(* IEC 61131-3 sources: plcassist-cli/packages/volt-lsp-iec/test-corpus/bakon-nano/Device/Plc Logic/Application/Library Manager/FloatingPointUtils, 43 files *)

(* ---- GVL.gvl ---- *)
VAR_GLOBAL
	EXP_MASK_REAL : UDINT := 16#7F800000;
	EXP_OFFSET_REAL : INT := 23;
	MANT_MASK_REAL : UDINT := 16#7FFFFF;
	RES_EXP_REAL : UINT := 16#FF;
	EXP_BIAS_REAL : INT := 127;
	NORM_MANT_REAL : UDINT := 16#800000;
	MAX_MANT_REAL : UDINT := 16#FFFFFF;
	MIN_EXP_REAL : INT := (INT#1 - (EXP_BIAS_REAL + EXP_OFFSET_REAL));
	MAX_EXP_REAL : INT := (UINT_TO_INT(RES_EXP_REAL) - ((INT#1 + EXP_BIAS_REAL) + EXP_OFFSET_REAL));
	EXP_MASK_LREAL : ULINT := 16#7FF0000000000000;
	EXP_OFFSET_LREAL : INT := 52;
	MANT_MASK_LREAL : ULINT := 16#FFFFFFFFFFFFF;
	RES_EXP_LREAL : UINT := 16#7FF;
	EXP_BIAS_LREAL : INT := 1023;
	NORM_MANT_LREAL : ULINT := 16#10000000000000;
	MAX_MANT_LREAL : ULINT := 16#1FFFFFFFFFFFFF;
	MIN_EXP_LREAL : INT := (INT#1 - (EXP_BIAS_LREAL + EXP_OFFSET_LREAL));
	MAX_EXP_LREAL : INT := (UINT_TO_INT(RES_EXP_LREAL) - ((INT#1 + EXP_BIAS_LREAL) + EXP_OFFSET_LREAL));
	STR_NAN : STRING(16) := 'NaN';
	STR_PINF : STRING(16) := '+Inf';
	STR_NINF : STRING(16) := '-Inf';
	LINT_MAX : LINT := 16#7FFFFFFFFFFFFFFF;
	INT_MAX : INT := 16#7FFF;
	INT_MIN : INT := -16#8000;
	DINT_MIN : DINT := -16#8000000;
	DINT_MAX : DINT := 16#7FFFFFFF;
END_VAR

(* ---- CEIL.fun ---- *)
FUNCTION CEIL : LREAL
VAR_INPUT
	F : LREAL;
END_VAR
END_FUNCTION

(* ---- CEILF.fun ---- *)
FUNCTION CEILF : REAL
VAR_INPUT
	F : REAL;
END_VAR
END_FUNCTION

(* ---- CHAREQCI.fun ---- *)
FUNCTION CHAREQCI : BOOL
VAR_INPUT
	C1 : BYTE;
	C2 : BYTE;
END_VAR
END_FUNCTION

(* ---- COMPOSELREAL.fun ---- *)
FUNCTION COMPOSELREAL : BOOL
VAR_INPUT
	LIM : LINT;
	IE : INT;
END_VAR
VAR_OUTPUT
	F : LREAL;
END_VAR
END_FUNCTION

(* ---- COMPOSELREALRAW.fun ---- *)
FUNCTION COMPOSELREALRAW : LREAL
VAR_INPUT
	BS : BOOL;
	UIE : UINT;
	ULIM : ULINT;
END_VAR
END_FUNCTION

(* ---- COMPOSEREAL.fun ---- *)
FUNCTION COMPOSEREAL : BOOL
VAR_INPUT
	DIM : DINT;
	IE : INT;
END_VAR
VAR_OUTPUT
	F : REAL;
END_VAR
END_FUNCTION

(* ---- COMPOSEREALRAW.fun ---- *)
FUNCTION COMPOSEREALRAW : REAL
VAR_INPUT
	BS : BOOL;
	UIE : UINT;
	UDIM : UDINT;
END_VAR
END_FUNCTION

(* ---- DESERIALIZEHEXREAL.fun ---- *)
FUNCTION DESERIALIZEHEXREAL : BOOL
VAR_INPUT
	PS : POINTER TO BYTE;
END_VAR
VAR_OUTPUT
	LIM : LINT;
	IE : INT;
	XNAN : BOOL;
	XINF : BOOL;
END_VAR
END_FUNCTION

(* ---- EXTRACTLREAL.fun ---- *)
FUNCTION EXTRACTLREAL : BOOL
VAR_INPUT
	F : LREAL;
END_VAR
VAR_OUTPUT
	IE : INT;
	LIM : LINT;
	XNAN : BOOL;
	XINF : BOOL;
END_VAR
END_FUNCTION

(* ---- EXTRACTLREALRAW.fun ---- *)
FUNCTION EXTRACTLREALRAW : BOOL
VAR_INPUT
	F : LREAL;
END_VAR
VAR_OUTPUT
	BS : BOOL;
	UIE : UINT;
	ULIM : ULINT;
END_VAR
END_FUNCTION

(* ---- EXTRACTREAL.fun ---- *)
FUNCTION EXTRACTREAL : BOOL
VAR_INPUT
	F : REAL;
END_VAR
VAR_OUTPUT
	IE : INT;
	DIM : DINT;
	XNAN : BOOL;
	XINF : BOOL;
END_VAR
END_FUNCTION

(* ---- EXTRACTREALRAW.fun ---- *)
FUNCTION EXTRACTREALRAW : BOOL
VAR_INPUT
	F : REAL;
END_VAR
VAR_OUTPUT
	BS : BOOL;
	UIE : UINT;
	UDIM : UDINT;
END_VAR
END_FUNCTION

(* ---- FLOOR.fun ---- *)
FUNCTION FLOOR : LREAL
VAR_INPUT
	F : LREAL;
END_VAR
END_FUNCTION

(* ---- FLOORF.fun ---- *)
FUNCTION FLOORF : REAL
VAR_INPUT
	F : REAL;
END_VAR
END_FUNCTION

(* ---- FLOORTEST.fun ---- *)
FUNCTION FLOORTEST : LREAL
VAR_INPUT
	F : LREAL;
END_VAR
END_FUNCTION

(* ---- GETLREALSPECIALVAL.fun ---- *)
FUNCTION GETLREALSPECIALVAL : LREAL
VAR_INPUT
	SV : ESpecial_FP_Value;
END_VAR
END_FUNCTION

(* ---- GETREALSPECIALVAL.fun ---- *)
FUNCTION GETREALSPECIALVAL : REAL
VAR_INPUT
	SV : ESpecial_FP_Value;
END_VAR
END_FUNCTION

(* ---- HEXDIGVAL.fun ---- *)
FUNCTION HEXDIGVAL : BYTE
VAR_INPUT
	C : BYTE;
END_VAR
END_FUNCTION

(* ---- HEXSTRTOLREAL.fun ---- *)
FUNCTION HEXSTRTOLREAL : BOOL
VAR_INPUT
	STR : STRING;
END_VAR
VAR_OUTPUT
	F : LREAL;
END_VAR
END_FUNCTION

(* ---- HEXSTRTOREAL.fun ---- *)
FUNCTION HEXSTRTOREAL : BOOL
VAR_INPUT
	STR : STRING;
END_VAR
VAR_OUTPUT
	F : REAL;
END_VAR
END_FUNCTION

(* ---- INSERTSTR.fun ---- *)
FUNCTION INSERTSTR : INT
VAR_INPUT
	PDST : POINTER TO BYTE;
	ISTARTINDEX : INT;
	PSRC : POINTER TO BYTE;
END_VAR
END_FUNCTION

(* ---- ISHEXDIG.fun ---- *)
FUNCTION ISHEXDIG : BOOL
VAR_INPUT
	C : BYTE;
END_VAR
END_FUNCTION

(* ---- ISLREALNAN.fun ---- *)
FUNCTION ISLREALNAN : BOOL
VAR_INPUT
	F : LREAL;
END_VAR
END_FUNCTION

(* ---- ISLREALNEGINFINITY.fun ---- *)
FUNCTION ISLREALNEGINFINITY : BOOL
VAR_INPUT
	F : LREAL;
END_VAR
END_FUNCTION

(* ---- ISLREALNUMBER.fun ---- *)
FUNCTION ISLREALNUMBER : BOOL
VAR_INPUT
	F : LREAL;
END_VAR
END_FUNCTION

(* ---- ISLREALPOSINFINITY.fun ---- *)
FUNCTION ISLREALPOSINFINITY : BOOL
VAR_INPUT
	F : LREAL;
END_VAR
END_FUNCTION

(* ---- ISREALNAN.fun ---- *)
FUNCTION ISREALNAN : BOOL
VAR_INPUT
	F : REAL;
END_VAR
END_FUNCTION

(* ---- ISREALNEGINFINITY.fun ---- *)
FUNCTION ISREALNEGINFINITY : BOOL
VAR_INPUT
	F : REAL;
END_VAR
END_FUNCTION

(* ---- ISREALNUMBER.fun ---- *)
FUNCTION ISREALNUMBER : BOOL
VAR_INPUT
	F : REAL;
END_VAR
END_FUNCTION

(* ---- ISREALPOSINFINITY.fun ---- *)
FUNCTION ISREALPOSINFINITY : BOOL
VAR_INPUT
	F : REAL;
END_VAR
END_FUNCTION

(* ---- LREALTOHEXSTR.fun ---- *)
FUNCTION LREALTOHEXSTR : STRING(32)
VAR_INPUT
	F : LREAL;
END_VAR
END_FUNCTION

(* ---- LREALTOSTR.fun ---- *)
FUNCTION LREALTOSTR : STRING(32)
VAR_INPUT
	F : LREAL;
END_VAR
END_FUNCTION

(* ---- REALTOHEXSTR.fun ---- *)
FUNCTION REALTOHEXSTR : STRING(32)
VAR_INPUT
	F : REAL;
END_VAR
END_FUNCTION

(* ---- REALTOSTR.fun ---- *)
FUNCTION REALTOSTR : STRING(16)
VAR_INPUT
	F : REAL;
END_VAR
END_FUNCTION

(* ---- SCANCONSTI.fun ---- *)
FUNCTION SCANCONSTI : BOOL
VAR_INPUT
	PS : POINTER TO BYTE;
	PSCONST : POINTER TO BYTE;
END_VAR
VAR_IN_OUT
	IDX : INT;
END_VAR
END_FUNCTION

(* ---- SCANHEXNUMERAL.fun ---- *)
FUNCTION SCANHEXNUMERAL : BOOL
VAR_INPUT
	PS : POINTER TO BYTE;
END_VAR
VAR_OUTPUT
	LI : LINT;
END_VAR
VAR_IN_OUT
	IDX : INT;
END_VAR
END_FUNCTION

(* ---- SERIALIZEHEXREAL.fun ---- *)
FUNCTION SERIALIZEHEXREAL : STRING(32)
VAR_INPUT
	LIM : LINT;
	IE : INT;
END_VAR
END_FUNCTION

(* ---- STRTOLREAL.fun ---- *)
FUNCTION STRTOLREAL : LREAL
VAR_INPUT
	STR : STRING;
END_VAR
END_FUNCTION

(* ---- STRTOREAL.fun ---- *)
FUNCTION STRTOREAL : REAL
VAR_INPUT
	STR : STRING;
END_VAR
END_FUNCTION

(* ---- TOHEXNUMERAL.fun ---- *)
FUNCTION TOHEXNUMERAL : INT
VAR_INPUT
	PDST : POINTER TO BYTE;
	LI : LINT;
END_VAR
END_FUNCTION

(* ---- TRUNCATE.fun ---- *)
FUNCTION TRUNCATE : LREAL
VAR_INPUT
	F : LREAL;
END_VAR
END_FUNCTION

(* ---- TRUNCATEF.fun ---- *)
FUNCTION TRUNCATEF : REAL
VAR_INPUT
	F : REAL;
END_VAR
END_FUNCTION
